(* IEC 61131-3 sources: stratumak/src/stmak/internal/modcompile/st/testdata/accept, 20 files *)

(* ---- actions.st ---- *)
{attribute 'summary' := 'Named pieces of a body, shared with it'}
{attribute 'license' := 'GPL'}

(* An ACTION is a named piece of a POU's body.  It shares every variable of the
   POU and has none of its own, which is what makes it different from a
   FUNCTION_BLOCK: nothing has to be passed in, and nothing has its own state.

   The alternative for splitting a long cyclic body is a function block, which
   changes the state layout and forces every touched variable through an
   interface, or a FUNCTION, which cannot see the POU's variables at all. *)

FUNCTION_BLOCK Counter
  VAR_INPUT
    step  : DINT;
    reset : BOOL;
  END_VAR
  VAR_OUTPUT
    total : DINT;
  END_VAR
  VAR
    overflows : DINT;
  END_VAR

  IF reset THEN
    clear();
  ELSE
    accumulate();
  END_IF;

(* An action of a function block reaches the instance, so its signature is the
   block body's exactly. *)
ACTION clear:
  total := 0;
  overflows := 0;
END_ACTION

ACTION accumulate:
  total := total + step;
  IF total > 1000 THEN
    overflows := overflows + 1;
    clear();
  END_IF;
END_ACTION

END_FUNCTION_BLOCK

{attribute 'doc' := 'Runs the counter and reports on it.'}
PROGRAM actions
  VAR_INPUT
    enable : BOOL;
    amount : DINT := 1;
  END_VAR
  VAR_OUTPUT
    count   : DINT;
    running : BOOL;
    idle    : BOOL;
  END_VAR
  VAR
    c        : Counter;
    selected : DINT;
  END_VAR

  (* An action of an instance, called from outside the block that declares
     it: `motor.stop()`.  It shares that instance's variables and takes no
     arguments -- there is no interface to pass anything through. *)
  c.clear();

  IF enable THEN
    (* An action of a PROGRAM sees the pin snapshot, so it may read and write
       pins exactly as the body does. *)
    advance(selected := amount);
  ELSE
    stop();
  END_IF;

  report();

ACTION advance:
  c(step := selected, reset := FALSE);
  count := c.total;
  running := TRUE;
END_ACTION

ACTION stop:
  c(step := 0, reset := TRUE);
  count := 0;
  running := FALSE;
END_ACTION

(* This one touches no pin at all, only instance state. *)
ACTION report:
  idle := NOT running;
END_ACTION

END_PROGRAM

(* ---- atmap.st ---- *)
{attribute 'summary' := 'Explicit pin mapping with AT'}
{attribute 'license' := 'GPL'}

(* A function block that publishes one of its own values to HAL.  It is not a
   VAR_INPUT, so nothing at a call site writes it -- the direction in the AT
   clause is the whole story, and there is no second writer to conflict with. *)

FUNCTION_BLOCK Axis
  VAR_INPUT
    cmd : LREAL;
  END_VAR
  VAR
    pos AT %Q.position : LREAL;
    err AT %Q.error    : LREAL;
    home AT %I.at_home : BOOL;
  END_VAR

  IF home THEN
    pos := 0.0;
  ELSE
    pos := pos + (cmd - pos) * 0.1;
  END_IF;
  err := cmd - pos;
END_FUNCTION_BLOCK

PROGRAM atmap
  VAR
    (* A plain VAR mapped explicitly, and renamed on the way out. *)
    enable  AT %I         : BOOL;
    running AT %Q.active  : BOOL;
    feed    AT %IO        : LREAL;

    x    : Axis;
    axes : ARRAY[0..2] OF Axis;
    i    : DINT;
  END_VAR

  running := enable;
  x(cmd := feed);
  FOR i := 0 TO 2 DO
    axes[i](cmd := feed);
  END_FOR;
END_PROGRAM

(* ---- constants.st ---- *)
{attribute 'summary' := 'Named constants as bounds, limits and labels'}
{attribute 'license' := 'GPL'}

(* Real ST names its bounds far more often than it writes them out, and a
   constant is only useful where the compiler can see its value: sizing an
   array, bounding a FOR, labelling a CASE arm.  A constant written as an
   expression counts too -- (24 * 60) is a value, not a computation. *)

TYPE
  Mode  : (OFF, MANUAL, AUTO);
  State : (OFF, RUNNING, FAULT);
END_TYPE

FUNCTION_BLOCK History
  VAR CONSTANT
    SLOTS       : DINT := 8;
    LAST_SLOT   : DINT := SLOTS - 1;
    WINDOW      : DINT := (2 * 4);
  END_VAR
  VAR_INPUT
    sample : LREAL;
  END_VAR
  VAR_OUTPUT
    mean : LREAL;
  END_VAR
  VAR
    (* An array of a block's own constant: the bound has to resolve while the
       rest of the block's declarations are still being read. *)
    slot  : ARRAY[0..LAST_SLOT] OF LREAL;
    total : LREAL;
    i     : DINT;
  END_VAR

  FOR i := 0 TO LAST_SLOT - 1 DO
    slot[i] := slot[i + 1];
  END_FOR;
  slot[LAST_SLOT] := sample;

  total := 0.0;
  FOR i := 0 TO LAST_SLOT DO
    total := total + slot[i];
  END_FOR;
  mean := total / WINDOW;
END_FUNCTION_BLOCK

PROGRAM constants
  VAR CONSTANT
    CHANNELS       : DINT := 4;
    MINUTES_PER_DAY : DINT := (24 * 60);
    SCALE          : LREAL := 1.0 / 5.0;
  END_VAR
  VAR_INPUT
    raw     : ARRAY[0..3] OF LREAL;
    request : DINT := 0;
  END_VAR
  VAR_OUTPUT
    average : LREAL;
    minutes : DINT;
    active  : BOOL;
  END_VAR
  VAR
    hist : History;
    mode : Mode  := Mode.OFF;
    step : State := State.OFF;
    sum  : LREAL;
    i    : DINT;
  END_VAR

  sum := 0.0;
  FOR i := 0 TO CHANNELS - 1 DO
    sum := sum + raw[i];
  END_FOR;
  average := sum * SCALE;
  minutes := MINUTES_PER_DAY;

  hist(sample := average);

  (* Both enumerations declare OFF, so an unqualified OFF would be ambiguous;
     the qualified form says which is meant. *)
  CASE request OF
    0: mode := Mode.OFF;
    1: mode := Mode.MANUAL;
    2: mode := Mode.AUTO;
  ELSE
    mode := Mode.OFF;
  END_CASE;

  IF mode = Mode.OFF THEN
    step := State.OFF;
  ELSE
    step := State.RUNNING;
  END_IF;

  active := step = State.RUNNING;
END_PROGRAM

(* ---- durations.st ---- *)
{attribute 'summary' := 'The TIME type: literals, arithmetic and conversions'}
{attribute 'license' := 'GPL'}

(* A duration is held as int64 nanoseconds -- what get_time() and a task's
   period already are.  It is not a number: it adds to and compares with
   another duration, scales by a count, and divides by another duration to give
   their ratio, and anything else is refused rather than guessed at.

   See docs/dev/MODCOMPILE_ST_STDLIB.md §5. *)

TYPE Config : STRUCT
  (* The shape the production sources actually use: PT is read from a struct
     member far more often than it is written as a literal. *)
  errDelay  : TIME;
  pumpOff   : TIME;
END_STRUCT
END_TYPE

FUNCTION_BLOCK Elapsed
  VAR_INPUT
    run : BOOL;
  END_VAR
  VAR_OUTPUT
    et : TIME;
  END_VAR

  IF run THEN
    (* fperiod is LREAL seconds, so the bridge is named for seconds. *)
    et := et + SECONDS_TO_TIME(fperiod);
  ELSE
    et := T#0s;
  END_IF;
END_FUNCTION_BLOCK

PROGRAM durations
  VAR_INPUT
    run : BOOL;
    (* HAL has no duration type, so a settable one arrives as seconds. *)
    delay_s : LREAL;
  END_VAR
  VAR_OUTPUT
    expired    : BOOL;
    elapsed_ms : DINT;
    remaining  : LREAL;
    fraction   : LREAL;
  END_VAR
  VAR
    cfg : Config;
    e   : Elapsed;

    pt      : TIME := T#500ms;
    warmup  : TIME := T#1m30s;
    fine    : TIME := T#1s500ms250us;
    half    : TIME;
  END_VAR

  cfg.errDelay := SECONDS_TO_TIME(delay_s);
  cfg.pumpOff  := T#2s;

  e(run := run);

  expired    := e.et >= pt;
  elapsed_ms := TIME_TO_DINT(e.et);
  remaining  := TIME_TO_SECONDS(warmup - e.et);
  fraction   := e.et / pt;

  (* Scaling: by a whole count and by a fraction. *)
  half := pt / 2;
  pt   := half * 2;
  warmup := warmup * 1.5;

  IF cfg.errDelay > cfg.pumpOff THEN
    pt := fine;
  END_IF;
END_PROGRAM

(* ---- fbnest.st ---- *)
{attribute 'summary' := 'Nested and arrayed function block instances'}
{attribute 'license' := 'GPL'}

(* A function block instance nests as a struct inside inst_t, so an FB may
   contain another, and an array of instances is unremarkable -- neither
   would be true if instances carried HAL identities of their own. *)

FUNCTION_BLOCK Accumulator
  VAR_INPUT
    add   : LREAL;
    clear : BOOL;
  END_VAR
  VAR_OUTPUT
    total : LREAL;
  END_VAR

  IF clear THEN
    total := 0.0;
  ELSE
    total := total + add;
  END_IF;
END_FUNCTION_BLOCK

FUNCTION_BLOCK Averager
  VAR_INPUT
    sample : LREAL;
    reset  : BOOL;
  END_VAR
  VAR_OUTPUT
    mean : LREAL;
  END_VAR
  VAR
    acc   : Accumulator;
    count : DINT;
  END_VAR

  IF reset THEN
    count := 0;
  ELSE
    count := count + 1;
  END_IF;

  acc(add := sample, clear := reset);

  IF count > 0 THEN
    mean := acc.total / count;
  ELSE
    mean := 0.0;
  END_IF;
END_FUNCTION_BLOCK

PROGRAM fbnest
  VAR_INPUT
    ch    : ARRAY[0..3] OF LREAL;
    reset : BOOL;
  END_VAR
  VAR_OUTPUT
    mean0 : LREAL;
    mean1 : LREAL;
  END_VAR
  VAR
    avg : ARRAY[0..3] OF Averager;
    i   : DINT;
  END_VAR

  FOR i := 0 TO 3 DO
    avg[i](sample := ch[i], reset := reset);
  END_FOR;

  mean0 := avg[0].mean;
  mean1 := avg[1].mean;
END_PROGRAM

(* ---- methods.st ---- *)
{attribute 'summary' := 'Methods on a function block instance'}
{attribute 'license' := 'GPL'}

(* A METHOD is an operation on an instance: it has its own interface and its
   own locals, and it can reach the instance's variables.  That is what makes
   it different from an ACTION, which shares the POU's variables and has no
   interface at all -- and why both can share the `inst.name()` call syntax
   without either having to know about the other.

   See docs/dev/MODCOMPILE_ST_STDLIB.md §7a. *)

FUNCTION_BLOCK Accumulator
  VAR_OUTPUT
    total : DINT;
  END_VAR
  VAR
    calls : DINT;
  END_VAR

  calls := calls + 1;

  (* The block's own body reaching one of its methods, IEC's way round. *)
  IF calls = 1 THEN
    THIS^.clear();
  END_IF;

{attribute 'doc' := 'Add a weighted value and report the new total.'}
METHOD add : DINT
  VAR_INPUT
    n      : DINT;
    weight : DINT;
  END_VAR
  VAR
    (* A method's own local, which does not persist between calls -- that is
       what the block's VAR is for. *)
    scaled : DINT;
  END_VAR

  scaled := n * weight;
  total  := total + scaled;
  add    := total;
END_METHOD

{attribute 'doc' := 'Add one, at the standard weight.'}
METHOD tick : DINT
  (* A sibling method, called with no name for the instance: there is one in
     scope either way, and the generated function already has it. *)
  tick := add(n := 1, weight := 1);
END_METHOD

{attribute 'doc' := 'Start again.'}
METHOD clear
  (* No result type at all: a method that only acts on the instance returns
     nothing, and writing `: VOID` for that would need a type ST does not
     have. *)
  total := 0;
END_METHOD

(* An action beside the methods, sharing the block's variables and taking no
   interface of its own. *)
ACTION note:
  calls := calls + 1;
END_ACTION

END_FUNCTION_BLOCK

PROGRAM methods
  VAR_INPUT
    reset : BOOL;
  END_VAR
  VAR_OUTPUT
    running : DINT;
  END_VAR
  VAR
    acc : Accumulator;
  END_VAR

  acc();

  (* As an expression, for the result... *)
  running := acc.add(n := 5, weight := 2);

  (* ...and as a statement, where there is none to use. *)
  IF reset THEN
    acc.clear();
  END_IF;

  (* The same spelling reaches an action, which is the point of §7a. *)
  acc.note();
END_PROGRAM

(* ---- params.st ---- *)
{attribute 'summary' := 'HAL parameters, at the top level and inside a block'}
{attribute 'license' := 'GPL'}

(* A HAL parameter is a value in shared memory that no signal connects to.
   `AT %MRW` is a tunable HAL sets and the component reads; `AT %MR` is a
   diagnostic the component writes and HAL only reads.  See §3.5. *)

FUNCTION_BLOCK Limiter
  VAR_INPUT
    raw : LREAL;
  END_VAR
  VAR_OUTPUT
    limited : LREAL;
  END_VAR
  VAR
    (* A parameter inside a block becomes one per instance, named by the
       path that reaches it -- exactly as a published pin is. *)
    ceiling AT %MRW        : LREAL := 100.0;
    hits    AT %MR.clamped : DINT;
  END_VAR

  limited := raw;
  IF limited > ceiling THEN
    limited := ceiling;
    hits := hits + 1;
  END_IF;
END_FUNCTION_BLOCK

PROGRAM params
  VAR_INPUT
    cmd : LREAL;
  END_VAR
  VAR_OUTPUT
    out : LREAL;
  END_VAR
  VAR
    {attribute 'doc' := 'Multiplies the command before limiting.'}
    gain    AT %MRW       : LREAL := 1.0;
    {attribute 'doc' := 'Set when the last cycle was scaled down.'}
    scaled  AT %MR.active : BOOL;
    invert  AT %MRW       : BOOL;

    lim : Limiter;
  END_VAR

  lim(raw := cmd * gain);
  out := lim.limited;
  IF invert THEN
    out := -out;
  END_IF;
  scaled := gain < 1.0;
END_PROGRAM

(* ---- period.st ---- *)
{attribute 'summary' := 'fperiod, in each kind of body that may use it'}
{attribute 'license' := 'GPL'}

(* fperiod is the period of the thread this body is running in.  The backend
   reaches it two ways -- from the HAL function's own argument where that is in
   scope, and from the RT task otherwise -- and they are the same number,
   because a HAL function is invoked by its own thread.  See
   docs/dev/MODCOMPILE_ST_STDLIB.md §4. *)

FUNCTION_BLOCK Integrator
  VAR_INPUT
    rate : LREAL;
  END_VAR
  VAR_OUTPUT
    total : LREAL;
  END_VAR

  (* A block body is its own C function and was never handed the argument. *)
  IF rate = 0.0 THEN
    reset();
  ELSE
    total := total + rate * fperiod;
  END_IF;

ACTION reset:
  total := 0.0;
END_ACTION

END_FUNCTION_BLOCK

PROGRAM period
  VAR_INPUT
    enable : BOOL;
    rate   : LREAL;
  END_VAR
  VAR_OUTPUT
    total   : LREAL;
    elapsed : LREAL;
  END_VAR
  VAR
    acc : Integrator;
  END_VAR

  IF enable THEN
    (* An exported body has the argument. *)
    elapsed := elapsed + fperiod;
    acc(rate := rate);
  ELSE
    stop();
  END_IF;
  total := acc.total;

(* An action is its own C function too, even inside a PROGRAM. *)
ACTION stop:
  elapsed := 0.0;
END_ACTION

END_PROGRAM

(* ---- ramplimit.st ---- *)
{attribute 'summary' := 'Rate-limited position follower'}
{attribute 'license' := 'GPL'}
{attribute 'author'  := 'stratuMAK'}

(* The worked example of docs/dev/MODCOMPILE_ST_FRONTEND.md §3.  A function
   block is internal: Ramp has no HAL identity, only ramplimit's own
   VAR_INPUT/VAR_OUTPUT become pins.  Where a sub-component's input should be
   wirable, declare the pin at PROGRAM level and pass it in -- which is what
   `target := target` does here. *)

FUNCTION_BLOCK Ramp
  VAR_INPUT
    target : LREAL;
    rate   : LREAL;
    dt     : LREAL;
  END_VAR
  VAR_OUTPUT
    out    : LREAL;
  END_VAR
  VAR
    step   : LREAL;
  END_VAR

  step := rate * dt;
  IF target > out + step THEN
    out := out + step;
  ELSIF target < out - step THEN
    out := out - step;
  ELSE
    out := target;
  END_IF;
END_FUNCTION_BLOCK

PROGRAM ramplimit
  VAR_INPUT
    {attribute 'doc' := 'Commanded position.'}
    target   : LREAL;
    {attribute 'doc' := 'Maximum rate of change, units per second.'}
    max_rate : LREAL := 10.0;
    enable   : BOOL;
  END_VAR
  VAR_OUTPUT
    out      : LREAL;
  END_VAR
  VAR
    r : Ramp;
  END_VAR

  IF enable THEN
    r(target := target, rate := max_rate, dt := fperiod);
    out := r.out;
  ELSE
    out := target;
  END_IF;
END_PROGRAM

(* ---- and2.st ---- *)
{attribute 'summary' := 'Two-input AND gate'}
{attribute 'license' := 'GPL'}
{attribute 'author'  := 'stratuMAK'}

(* The smallest useful component: two inputs, one output, no state.
   The .comp equivalent is src/hal/components/and2.comp. *)

PROGRAM and2
  VAR_INPUT
    {attribute 'doc' := 'First input.'}
    in0 : BOOL;
    {attribute 'doc' := 'Second input.'}
    in1 : BOOL;
  END_VAR
  VAR_OUTPUT
    {attribute 'doc' := 'TRUE when both inputs are TRUE.'}
    out : BOOL;
  END_VAR

  out := in0 AND in1;
END_PROGRAM

(* ---- arrays.st ---- *)
{attribute 'summary' := 'Select and average from an array pin'}
{attribute 'license' := 'GPL'}

(* Array pins map one dimension only, since a HAL pin name carries one
   index: channel.0 .. channel.7.  Multi-dimensional arrays are fine as
   internal state.  The non-zero lower bound on `window` is deliberate --
   every index site has to subtract it. *)

PROGRAM arrays
  VAR_INPUT
    channel  : ARRAY[0..7] OF LREAL;
    selected : DINT := 0;
  END_VAR
  VAR_OUTPUT
    value   : LREAL;
    average : LREAL;
  END_VAR
  VAR
    window : ARRAY[1..4] OF LREAL;
    grid   : ARRAY[0..1, 0..2] OF LREAL;
    total  : LREAL;
    i, j   : DINT;
  END_VAR

  value := channel[selected];

  total := 0.0;
  FOR i := 0 TO 7 DO
    total := total + channel[i];
  END_FOR;
  average := total / 8.0;

  FOR i := 1 TO 4 DO
    window[i] := average;
  END_FOR;

  FOR i := 0 TO 1 DO
    FOR j := 0 TO 2 DO
      grid[i, j] := average;
    END_FOR;
  END_FOR;
END_PROGRAM

(* ---- documented.st ---- *)
{attribute 'summary'     := 'Every documentation field, exercised'}
{attribute 'description' := 'A component that exists to prove its man page is as complete as one generated from a .comp: description, function docs, per-pin docs, notes, examples, author, licence and see-also.'}
{attribute 'license'     := 'GPL'}
{attribute 'author'      := 'stratuMAK'}
{attribute 'see_also'    := '\fBscale\fR(9), \fBand2\fR(9).'}
{attribute 'notes'       := 'The two functions may run in different threads; only \fBupdate\fR needs a floating-point one.'}
{attribute 'examples'    := 'loadrt documented$Naddf documented.sample servo-thread$Naddf documented.update servo-thread'}

(* Metadata before the first declaration describes the component.  A pragma
   heading a PROGRAM documents that program's HAL function, and one inside a
   VAR section documents the pin it precedes. *)

VAR_GLOBAL
  latest : DINT;
END_VAR

{attribute 'doc' := 'Latches the raw input when strobed. Uses no floating point.'}
PROGRAM sample
  VAR_INPUT
    {attribute 'doc' := 'Value to latch.'}
    raw : DINT;
    {attribute 'doc' := 'Rising level latches \fBraw\fR.'}
    strobe : BOOL;
  END_VAR
  VAR_OUTPUT
    {attribute 'doc' := 'TRUE once a value has been latched.'}
    valid : BOOL;
  END_VAR

  IF strobe THEN
    latest := raw;
    valid := TRUE;
  END_IF;
END_PROGRAM

{attribute 'doc' := 'Scales the latched value. Requires a floating-point thread.'}
PROGRAM update
  VAR_INPUT
    {attribute 'doc' := 'Multiplier applied to the latched value.'}
    gain : LREAL := 1.0;
  END_VAR
  VAR_OUTPUT
    {attribute 'doc' := 'The latched value times \fBgain\fR.'}
    scaled : LREAL;
  END_VAR

  scaled := latest * gain;
END_PROGRAM

(* ---- funcs.st ---- *)
{attribute 'summary' := 'Stateless helper functions'}
{attribute 'license' := 'GPL'}

(* A FUNCTION keeps no state between calls, so it may be called from an
   expression -- unlike a FUNCTION_BLOCK, whose invocation is a statement
   because it mutates its instance. *)

FUNCTION Clamp : LREAL
  VAR_INPUT
    value : LREAL;
    low   : LREAL;
    high  : LREAL;
  END_VAR

  IF value < low THEN
    Clamp := low;
  ELSIF value > high THEN
    Clamp := high;
  ELSE
    Clamp := value;
  END_IF;
END_FUNCTION

FUNCTION Lerp : LREAL
  VAR_INPUT
    a, b : LREAL;
    t    : LREAL;
  END_VAR
  VAR
    span : LREAL;
  END_VAR

  span := b - a;
  Lerp := a + span * Clamp(t, 0.0, 1.0);
END_FUNCTION

PROGRAM funcs
  VAR_INPUT
    raw  : LREAL;
    blend : LREAL;
  END_VAR
  VAR_OUTPUT
    limited : LREAL;
    mixed   : LREAL;
  END_VAR

  limited := Clamp(raw, -10.0, 10.0);
  mixed := Lerp(0.0, limited, blend);
END_PROGRAM

(* ---- literals.st ---- *)
{attribute 'summary' := 'Literal forms and operator precedence'}
{attribute 'license' := 'GPL'}

(* Spelled out because these are where a hand-written parser goes wrong
   quietly: based literals, digit separators, typed literals, and the
   precedence chain from ** down to OR. *)

PROGRAM literals
  VAR_INPUT
    enable : BOOL;
  END_VAR
  VAR_OUTPUT
    mask    : UDINT;
    result  : LREAL;
    decided : BOOL;
  END_VAR
  VAR
    a : DINT := 16#FF;
    b : DINT := 2#1010_1010;
    c : DINT := 8#777;
    d : DINT := 1_000_000;
    e : LREAL := 1.5;
    f : LREAL := 1.0E-3;
    g : LREAL := 2.5E3;
  END_VAR

  mask := UDINT#16#DEAD_BEEF;

  (* ** is right-associative and binds tighter than *; unary minus binds
     looser than ** on its left operand. *)
  result := e + f * g - 2.0 ** 3.0 ** 2.0;
  result := -result;
  result := (e + f) * g;

  (* MOD sits with * and /; comparison is looser than arithmetic; then
     equality, AND, XOR, OR. *)
  decided := a + 1 < b AND c MOD 8 = 7 OR NOT enable;
  decided := decided XOR (a > b);
  decided := enable & decided;
END_PROGRAM

(* ---- loops.st ---- *)
{attribute 'summary' := 'Bounded iteration'}
{attribute 'license' := 'GPL'}

(* Every loop in a HAL function body carries a bound the compiler can see.
   FOR is bounded by construction.  WHILE and REPEAT are not, so each needs
   an explicit max_iterations cap -- without one, sema rejects the statement.
   See docs/dev/MODCOMPILE_ST_FRONTEND.md §4. *)

PROGRAM loops
  VAR_INPUT
    target    : LREAL;
    tolerance : LREAL := 0.001;
  END_VAR
  VAR_OUTPUT
    estimate   : LREAL;
    iterations : DINT;
  END_VAR
  VAR
    guess : LREAL;
    i     : DINT;
  END_VAR

  guess := target / 2.0;
  iterations := 0;

  (* Newton-Raphson for a square root: iterative settling is a real pattern,
     and a bounded WHILE says so more honestly than a FOR with a break. *)
  {attribute 'max_iterations' := '50'}
  WHILE guess * guess - target > tolerance DO
    guess := (guess + target / guess) / 2.0;
    iterations := iterations + 1;
  END_WHILE;

  {attribute 'max_iterations' := '10'}
  REPEAT
    iterations := iterations + 1;
  UNTIL iterations > 5
  END_REPEAT;

  FOR i := 0 TO 9 DO
    IF i > 4 THEN
      EXIT;
    END_IF;
    iterations := iterations + 1;
  END_FOR;

  estimate := guess;
END_PROGRAM

(* ---- scale.st ---- *)
{attribute 'summary'     := 'Scale and offset a value'}
{attribute 'description' := 'Computes out := in * gain + offset, with the result clamped to [min, max] when limiting is enabled.'}
{attribute 'license'     := 'GPL'}
{attribute 'author'      := 'stratuMAK'}
{attribute 'see_also'    := '\fBmult2\fR(9), \fBsum2\fR(9).'}

(* Exercises the full metadata vocabulary docgen needs, plus LREAL
   arithmetic and an underscore name that becomes a hyphenated pin:
   max_limit here is mycomp.max-limit in HAL. *)

PROGRAM scale
  VAR_INPUT
    in        : LREAL;
    gain      : LREAL := 1.0;
    offset    : LREAL := 0.0;
    limiting  : BOOL;
    min_limit : LREAL := -1.0E6;
    max_limit : LREAL := 1.0E6;
  END_VAR
  VAR_OUTPUT
    out       : LREAL;
    clamped   : BOOL;
  END_VAR
  VAR
    raw : LREAL;
  END_VAR

  raw := in * gain + offset;
  clamped := FALSE;

  IF limiting THEN
    IF raw > max_limit THEN
      raw := max_limit;
      clamped := TRUE;
    ELSIF raw < min_limit THEN
      raw := min_limit;
      clamped := TRUE;
    END_IF;
  END_IF;

  out := raw;
END_PROGRAM

(* ---- statemachine.st ---- *)
{attribute 'summary' := 'Three-state sequencer with a fault path'}
{attribute 'license' := 'GPL'}

(* An enumeration used as a state variable, with CASE arms labelled by
   constant name rather than by number.  Resolving those names is exactly
   what the standalone prototype could not do. *)

TYPE
  State : (IDLE, RUNNING, FAULTED);
END_TYPE

PROGRAM statemachine
  VAR_INPUT
    start   : BOOL;
    stop    : BOOL;
    fault   : BOOL;
    reset   : BOOL;
  END_VAR
  VAR_OUTPUT
    is_running : BOOL;
    alarm   : BOOL;
  END_VAR
  VAR
    state : State := IDLE;
  END_VAR

  IF fault THEN
    state := FAULTED;
  END_IF;

  CASE state OF
    IDLE:
      IF start AND NOT stop THEN
        state := RUNNING;
      END_IF;
    RUNNING:
      IF stop THEN
        state := IDLE;
      END_IF;
    FAULTED:
      IF reset AND NOT fault THEN
        state := IDLE;
      END_IF;
  ELSE
    state := FAULTED;
  END_CASE;

  is_running := state = RUNNING;
  alarm   := state = FAULTED;
END_PROGRAM

(* ---- structs.st ---- *)
{attribute 'summary' := 'Nested structures and indexed field assignment'}
{attribute 'license' := 'GPL'}

(* `pts[i].x := ...` is the lvalue shape the standalone prototype could not
   express at all: its assignment target was a name plus optional indices,
   not an expression. *)

TYPE
  Point : STRUCT
    x : LREAL;
    y : LREAL;
  END_STRUCT;

  Rect : STRUCT
    topLeft     : Point;
    bottomRight : Point;
  END_STRUCT;
END_TYPE

PROGRAM structs
  VAR_INPUT
    px    : LREAL;
    py    : LREAL;
    index : DINT := 0;
  END_VAR
  VAR_OUTPUT
    width  : LREAL;
    height : LREAL;
  END_VAR
  VAR
    cursor : Point;
    bounds : Rect;
    pts    : ARRAY[0..3] OF Point;
    i      : DINT;
  END_VAR

  cursor.x := px;
  cursor.y := py;

  pts[index].x := cursor.x;
  pts[index].y := cursor.y;

  bounds.topLeft.x := pts[0].x;
  bounds.topLeft.y := pts[0].y;
  bounds.bottomRight.x := pts[0].x;
  bounds.bottomRight.y := pts[0].y;

  FOR i := 1 TO 3 DO
    IF pts[i].x < bounds.topLeft.x THEN
      bounds.topLeft.x := pts[i].x;
    END_IF;
    IF pts[i].x > bounds.bottomRight.x THEN
      bounds.bottomRight.x := pts[i].x;
    END_IF;
  END_FOR;

  width  := bounds.bottomRight.x - bounds.topLeft.x;
  height := bounds.bottomRight.y - bounds.topLeft.y;
END_PROGRAM

(* ---- twoprograms.st ---- *)
{attribute 'summary' := 'Two thread functions sharing state'}
{attribute 'license' := 'GPL'}

(* One PROGRAM per exported HAL function.  These become twoprograms.read and
   twoprograms.write, addf-able to different threads, with VAR_GLOBAL the
   state they share.  Each PROGRAM carries its own pins.

   `read` touches no floating point, so it should export with fp = 0. *)

VAR_GLOBAL
  latched : DINT;
  ready   : BOOL;
END_VAR

PROGRAM read
  VAR_INPUT
    raw    : DINT;
    strobe : BOOL;
  END_VAR
  VAR_OUTPUT
    accepted : BOOL;
  END_VAR

  IF strobe THEN
    latched := raw;
    ready := TRUE;
  END_IF;
  accepted := ready;
END_PROGRAM

PROGRAM write
  VAR_INPUT
    gain : LREAL := 1.0;
  END_VAR
  VAR_OUTPUT
    scaled : LREAL;
    valid  : BOOL;
  END_VAR

  IF ready THEN
    scaled := latched * gain;
    valid  := TRUE;
  ELSE
    scaled := 0.0;
    valid  := FALSE;
  END_IF;
END_PROGRAM

(* ---- types.st ---- *)
{attribute 'summary' := 'Every type that reaches a HAL pin'}
{attribute 'license' := 'GPL'}

(* The pin side of the type table in docs/dev/MODCOMPILE_ST_FRONTEND.md §3.1.
   BOOL, DINT, UDINT and LREAL map exactly; SINT/INT and USINT/UINT are
   widened.  LINT, ULINT, TIME, STRING, STRUCT and FUNCTION_BLOCK cannot
   appear on a pin and stay internal here.  REAL on a pin is accepted with a
   warning, not rejected -- see reject/ for what is refused outright. *)

TYPE
  Celsius : LREAL;
  Counter : UDINT;
END_TYPE

PROGRAM types
  VAR_INPUT
    flag     : BOOL;
    small    : SINT;
    medium   : INT;
    large    : DINT;
    usmall   : USINT;
    umedium  : UINT;
    ularge   : UDINT;
    precise  : LREAL;
    temp     : Celsius;
    ticks    : Counter;
  END_VAR
  VAR_OUTPUT
    ok       : BOOL;
    sum      : DINT;
    scaled   : LREAL;
    ticked   : UDINT;
    widened  : UDINT;
  END_VAR
  VAR
    (* No HAL representation: internal only. *)
    wide     : LINT;
    uwide    : ULINT;
    label    : STRING[32];
    shortstr : STRING;
    approx   : REAL;
  END_VAR

  ok := flag;
  sum := small + medium + large;
  scaled := precise + temp;
  ticked := ticks + 1;
  wide := large;
  uwide := ularge;
  approx := 1.5;
  widened := ularge + usmall + umedium;
END_PROGRAM
